// TwinCAT 3 PLC project PLC
// ProgramVersion: 3.1.4026.16
// libraries:
//   Tc2_Standard, * (Beckhoff Automation GmbH)
//   Tc2_System, * (Beckhoff Automation GmbH)
// project tree:
//   GVLs/ GVL.TcGVL
//   / PlcTask.TcTTO
//   POUs/ MAIN.TcPOU
// real-time tasks:
//   TASK PlcTask: cycle T#10ms, priority 20, ADS port 350
// I/O:
//   DEVICE Device 1 (NOV-DP-RAM)
//   DEVICE Device 2 (Onboard I/O Device), AmsNetId 5.174.170.138.3.1
//     Term 1 (CX7028) [CX7028-0000-0121]
//       modules: Module 1 (DIO_2x), Module 2 (Empty Module), Module 3 (DIO_2x), Module 4 (Empty Module), Module 5 (DI_2x), Module 6 (Empty Module), Module 7 (DI_2x), Module 8 (Empty Module)
// variable links:
//   PLC/PLC Instance <-> Device 2 (Onboard I/O Device)/Term 1 (CX7028)
//     PlcTask Inputs/GVL.bEStopPressed <-> Module 1 (DIO_2x)/DIO_2x Input Channel 1/Input
//     PlcTask Inputs/GVL.bEStopPressed2 <-> Module 5 (DI_2x)/DI_2x Input Channel 1/Input
//     PlcTask Inputs/GVL.bEStopPressed3 <-> Module 7 (DI_2x)/DI_2x Input Channel 1/Input
//     PlcTask Inputs/GVL.bEStopPressed4 <-> Module 5 (DI_2x)/DI_2x Input Channel 2/Input
//     PlcTask Outputs/MAIN.xOUput1 <-> Module 1 (DIO_2x)/DIO_2x Output Channel 1/Output
//     PlcTask Outputs/MAIN.xOUput2 <-> Module 1 (DIO_2x)/DIO_2x Output Channel 2/Output
//     PlcTask Outputs/MAIN.xOUput3 <-> Module 3 (DIO_2x)/DIO_2x Output Channel 1/Output
//     PlcTask Outputs/MAIN.xOUput4 <-> Module 3 (DIO_2x)/DIO_2x Output Channel 2/Output

CONFIGURATION PLC
    RESOURCE PLC ON TwinCAT3
        TASK PlcTask(INTERVAL := T#10ms, PRIORITY := 20);
        PROGRAM MAIN WITH PlcTask : MAIN;
    END_RESOURCE
END_CONFIGURATION

// ---- GVLs/GVL.TcGVL
{attribute 'qualified_only'}
VAR_GLOBAL
		iCounter : INT;
		bEStopPressed AT %I* : BOOL;
		bEStopPressed2 AT %I* : BOOL;
		bEStopPressed3 AT %I* : BOOL;
		bEStopPressed4 AT %I* : BOOL;
END_VAR

// ---- POUs/MAIN.TcPOU
PROGRAM MAIN
VAR
iCase : INT := 0;
xOUput1 AT %Q* : BOOL;
xOUput2 AT %Q* : BOOL;
xOUput3 AT %Q* : BOOL;
xOUput4 AT %Q* : BOOL;
timetime : TON ;
END_VAR

WHILE GVL.bEStopPressed DO
GVL.iCounter := GVL.iCounter + 1;
END_WHILE



CASE iCase OF  
	0: 
	IF GVL.iCounter < 10 THEN
		xOUput1 := TRUE;
	END_IF
	
		IF GVL.iCounter > 10 AND GVL.iCounter < 30  THEN
		xOUput2 := TRUE;
	END_IF

	IF GVL.iCounter > 30 AND GVL.iCounter < 100  THEN
		xOUput3 := TRUE;
	END_IF
	IF  GVL.iCounter = 100 THEN
		iCase := 1;
	END_IF

	1: GVL.iCounter := GVL.iCounter - 1;
		IF GVL.iCounter < 10 THEN
		xOUput3 := FALSE;
	END_IF
	
		IF GVL.iCounter > 10 AND GVL.iCounter < 30  THEN
		xOUput2 := FALSE;
	END_IF

	IF GVL.iCounter > 30 AND GVL.iCounter < 100  THEN
		xOUput1 := FALSE;
	END_IF
	IF  GVL.iCounter = 0 THEN
		iCase := 0;
	END_IF

END_CASE

END_PROGRAM
